PROGRAM MAIN
VAR
    bManualMode AT %I* : BOOL;
    bRotateLeft AT %I* : BOOL;
    bRotateRight AT %I* : BOOL;
    bExtend AT %I* : BOOL;
    bRetract AT %I* : BOOL;
    bShift AT %I* : BOOL;
    bStopButton AT %I* : BOOL;

    bRotateLimit AT %I* : BOOL;
    bExtendLimit AT %I* : BOOL;
    bLiftLimit AT %I* : BOOL;
    bGripLimit AT %I* : BOOL;
	
	bAllButtonsReleased : BOOL;
	bShiftSelected : BOOL;
	bShiftMismatch : BOOL;
	bCommandArmed : BOOL;
	bMotionEnabled : BOOL;

    bRotateLeftCmd : BOOL;
    bRotateRightCmd : BOOL;
    bExtendCmd : BOOL;
    bRetractCmd : BOOL;
    bLiftUp : BOOL;
    bLiftDown : BOOL;
    bGripOpen : BOOL;
    bGripClose : BOOL;

    bReqRotateForward : BOOL;
    bReqRotateBackward : BOOL;
    bReqExtendForward : BOOL;
    bReqExtendBackward : BOOL;
    bReqLiftForward : BOOL;
    bReqLiftBackward : BOOL;
    bReqGripForward : BOOL;
    bReqGripBackward : BOOL;

    bRotateRun AT %Q* : BOOL;
    bRotateDirection AT %Q* : BOOL;

    bExtendRun AT %Q* : BOOL;
    bExtendDirection AT %Q* : BOOL;

    bLiftRun AT %Q* : BOOL;
    bLiftDirection AT %Q* : BOOL;

    bGripRun AT %Q* : BOOL;
    bGripDirection AT %Q* : BOOL;


    fbRotateSelector : FB_CommandSelector;
    fbExtendSelector : FB_CommandSelector;
    fbLiftSelector : FB_CommandSelector;
    fbGripSelector : FB_CommandSelector;

    fbRotateMotor : FB_MotorControl;
    fbExtendMotor : FB_MotorControl;
    fbLiftMotor : FB_MotorControl;
    fbGripMotor : FB_MotorControl;
	
	nSelectedMotor : INT := 0;
END_VAR

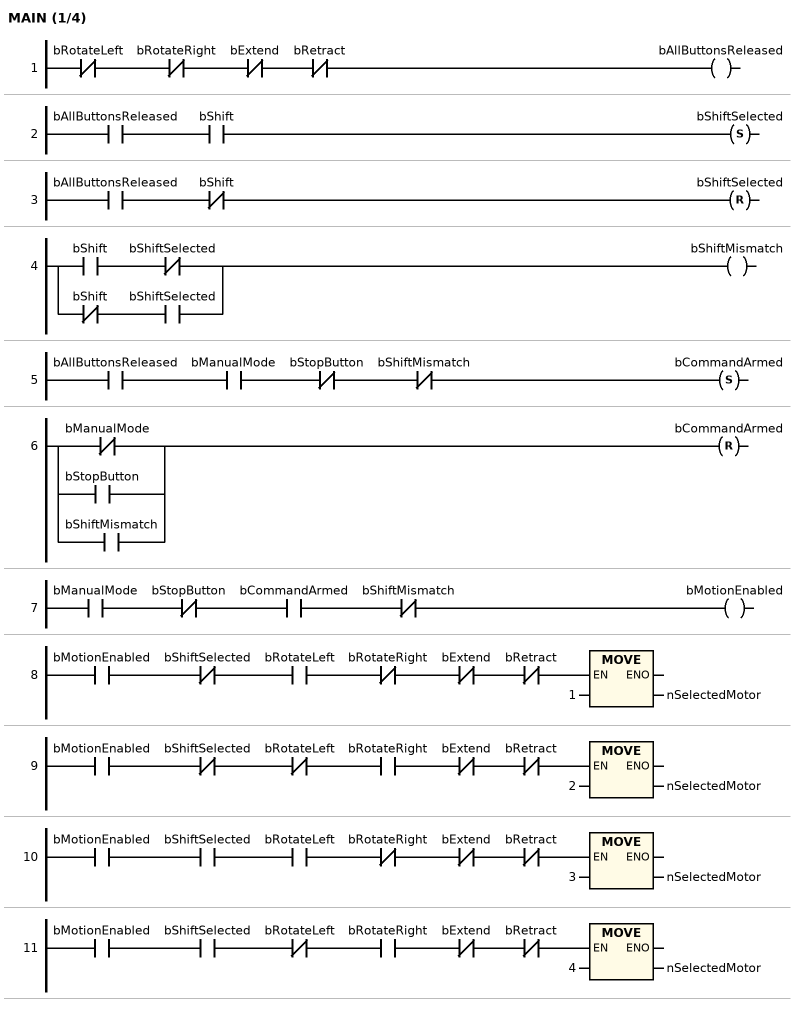
// NETWORK 1
bAllButtonsReleased := NOT bRotateLeft AND NOT bRotateRight AND NOT bExtend AND NOT bRetract;

// NETWORK 2
bShiftSelected S= bAllButtonsReleased AND bShift;

// NETWORK 3
bShiftSelected R= bAllButtonsReleased AND NOT bShift;

// NETWORK 4
bShiftMismatch := bShift AND NOT bShiftSelected OR NOT bShift AND bShiftSelected;

// NETWORK 5
bCommandArmed S= bAllButtonsReleased AND bManualMode AND NOT bStopButton AND NOT bShiftMismatch;

// NETWORK 6
bCommandArmed R= NOT bManualMode OR bStopButton OR bShiftMismatch;

// NETWORK 7
bMotionEnabled := bManualMode AND NOT bStopButton AND bCommandArmed AND NOT bShiftMismatch;

// NETWORK 8
IF bMotionEnabled AND NOT bShiftSelected AND bRotateLeft AND NOT bRotateRight AND NOT bExtend AND NOT bRetract THEN
    nSelectedMotor := 1;
END_IF

// NETWORK 9
IF bMotionEnabled AND NOT bShiftSelected AND NOT bRotateLeft AND bRotateRight AND NOT bExtend AND NOT bRetract THEN
    nSelectedMotor := 2;
END_IF

// NETWORK 10
IF bMotionEnabled AND bShiftSelected AND bRotateLeft AND NOT bRotateRight AND NOT bExtend AND NOT bRetract THEN
    nSelectedMotor := 3;
END_IF

// NETWORK 11
IF bMotionEnabled AND bShiftSelected AND NOT bRotateLeft AND bRotateRight AND NOT bExtend AND NOT bRetract THEN
    nSelectedMotor := 4;
END_IF

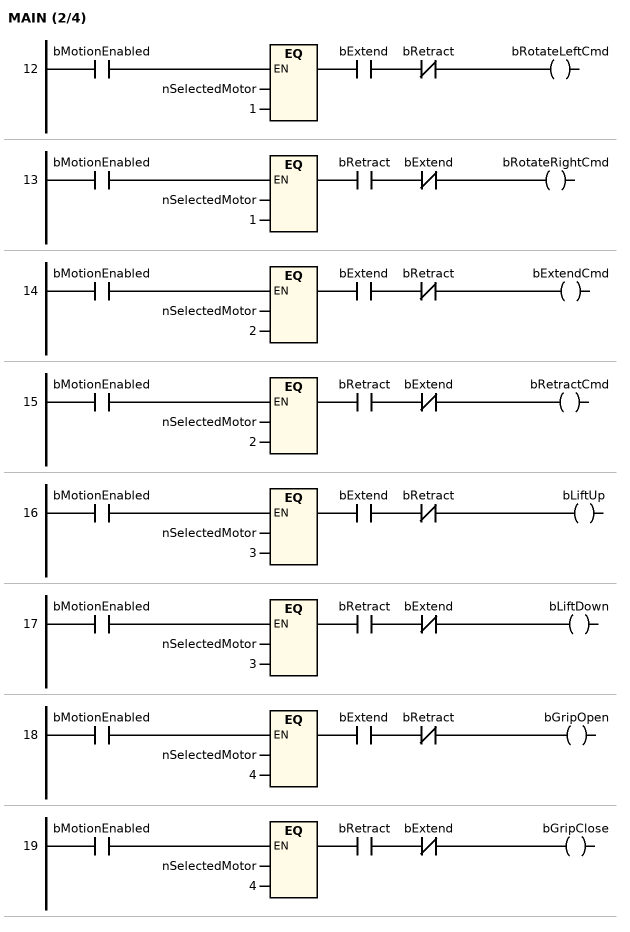
// NETWORK 12
bRotateLeftCmd := (bMotionEnabled AND nSelectedMotor = 1) AND bExtend AND NOT bRetract;

// NETWORK 13
bRotateRightCmd := (bMotionEnabled AND nSelectedMotor = 1) AND bRetract AND NOT bExtend;

// NETWORK 14
bExtendCmd := (bMotionEnabled AND nSelectedMotor = 2) AND bExtend AND NOT bRetract;

// NETWORK 15
bRetractCmd := (bMotionEnabled AND nSelectedMotor = 2) AND bRetract AND NOT bExtend;

// NETWORK 16
bLiftUp := (bMotionEnabled AND nSelectedMotor = 3) AND bExtend AND NOT bRetract;

// NETWORK 17
bLiftDown := (bMotionEnabled AND nSelectedMotor = 3) AND bRetract AND NOT bExtend;

// NETWORK 18
bGripOpen := (bMotionEnabled AND nSelectedMotor = 4) AND bExtend AND NOT bRetract;

// NETWORK 19
bGripClose := (bMotionEnabled AND nSelectedMotor = 4) AND bRetract AND NOT bExtend;

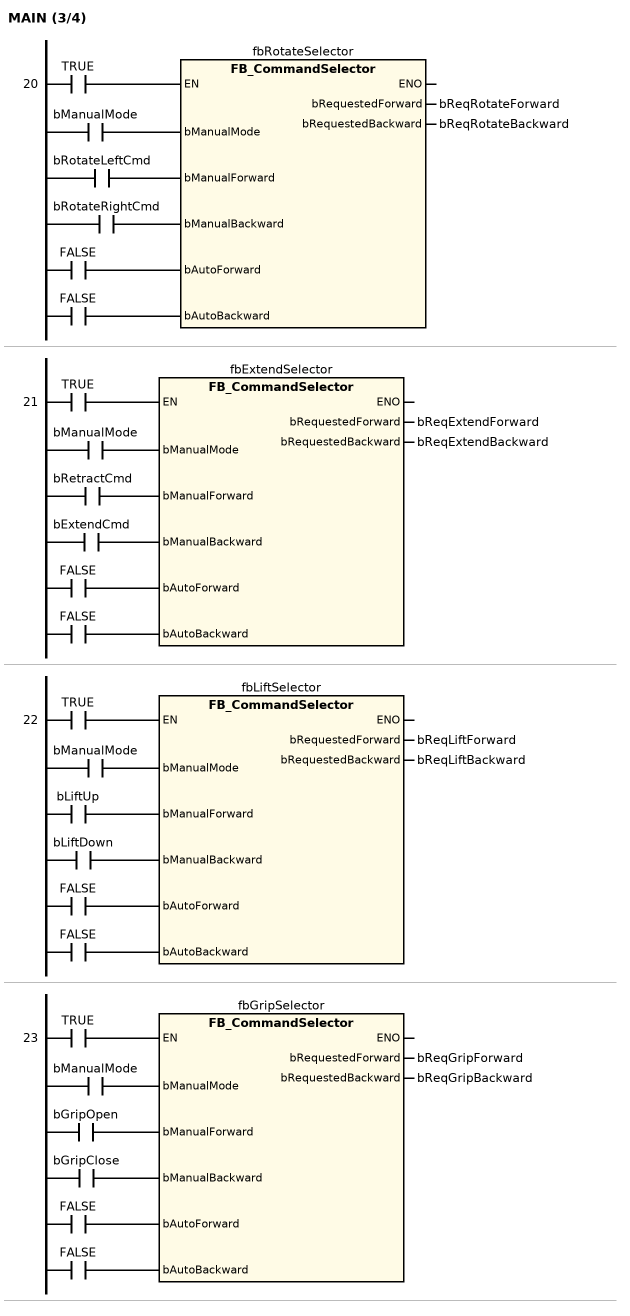
// NETWORK 20
fbRotateSelector(
    bManualMode := bManualMode,
    bManualForward := bRotateLeftCmd,
    bManualBackward := bRotateRightCmd,
    bAutoForward := FALSE,
    bAutoBackward := FALSE,
    bRequestedForward => bReqRotateForward,
    bRequestedBackward => bReqRotateBackward); // FB_CommandSelector

// NETWORK 21
fbExtendSelector(
    bManualMode := bManualMode,
    bManualForward := bRetractCmd,
    bManualBackward := bExtendCmd,
    bAutoForward := FALSE,
    bAutoBackward := FALSE,
    bRequestedForward => bReqExtendForward,
    bRequestedBackward => bReqExtendBackward); // FB_CommandSelector

// NETWORK 22
fbLiftSelector(
    bManualMode := bManualMode,
    bManualForward := bLiftUp,
    bManualBackward := bLiftDown,
    bAutoForward := FALSE,
    bAutoBackward := FALSE,
    bRequestedForward => bReqLiftForward,
    bRequestedBackward => bReqLiftBackward); // FB_CommandSelector

// NETWORK 23
fbGripSelector(
    bManualMode := bManualMode,
    bManualForward := bGripOpen,
    bManualBackward := bGripClose,
    bAutoForward := FALSE,
    bAutoBackward := FALSE,
    bRequestedForward => bReqGripForward,
    bRequestedBackward => bReqGripBackward); // FB_CommandSelector

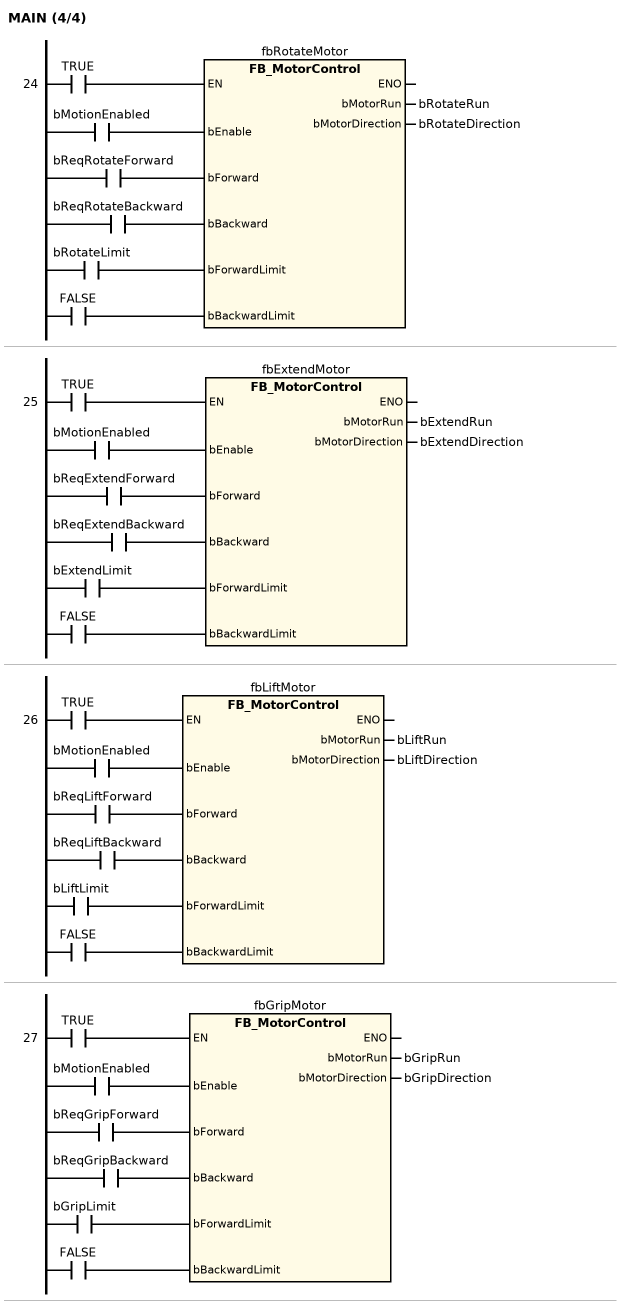
// NETWORK 24
fbRotateMotor(
    bEnable := bMotionEnabled,
    bForward := bReqRotateForward,
    bBackward := bReqRotateBackward,
    bForwardLimit := bRotateLimit,
    bBackwardLimit := FALSE,
    bMotorRun => bRotateRun,
    bMotorDirection => bRotateDirection); // FB_MotorControl

// NETWORK 25
fbExtendMotor(
    bEnable := bMotionEnabled,
    bForward := bReqExtendForward,
    bBackward := bReqExtendBackward,
    bForwardLimit := bExtendLimit,
    bBackwardLimit := FALSE,
    bMotorRun => bExtendRun,
    bMotorDirection => bExtendDirection); // FB_MotorControl

// NETWORK 26
fbLiftMotor(
    bEnable := bMotionEnabled,
    bForward := bReqLiftForward,
    bBackward := bReqLiftBackward,
    bForwardLimit := bLiftLimit,
    bBackwardLimit := FALSE,
    bMotorRun => bLiftRun,
    bMotorDirection => bLiftDirection); // FB_MotorControl

// NETWORK 27
fbGripMotor(
    bEnable := bMotionEnabled,
    bForward := bReqGripForward,
    bBackward := bReqGripBackward,
    bForwardLimit := bGripLimit,
    bBackwardLimit := FALSE,
    bMotorRun => bGripRun,
    bMotorDirection => bGripDirection); // FB_MotorControl

END_PROGRAM

(* stored: Version 1.1.0.1
   POU MAIN: Id {26f6676c-871c-4b33-aa99-0c46ab4a81a1}, SpecialFunc None *)
